TYPE "FRK_SetPayload"
VERSION : 0.1
   STRUCT
      Info { ExternalAccessible := 'False'; ExternalVisible := 'False'; ExternalWritable := 'False'} : "ST_ConfigSetInfo";
      Records { ExternalAccessible := 'False'; ExternalVisible := 'False'; ExternalWritable := 'False'} : Array[1..30] of "ST_ConfigRecord";
   END_STRUCT;

END_TYPE

